FUNCTION_BLOCK PID_DEMO_PROCESS (* Offline prototype; see docs/pid/README.md; native validation pending *)
  (* Standard: 61499-2 *)
  (* Version 0.1, 2026-10-18, Guilherme *)
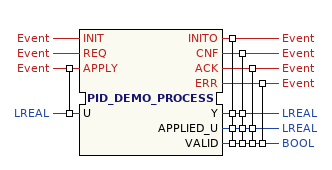
  EVENT_INPUT
    INIT;
    REQ;
    APPLY WITH U;
  END_EVENT
  EVENT_OUTPUT
    INITO WITH Y, APPLIED_U, VALID;
    CNF WITH Y, APPLIED_U, VALID;
    ACK WITH APPLIED_U, VALID;
    ERR WITH VALID;
  END_EVENT
  VAR_INPUT
    U : LREAL;
  END_VAR
  VAR_OUTPUT
    Y : LREAL;
    APPLIED_U : LREAL;
    VALID : BOOL;
  END_VAR
  VAR
    Y_NEXT : LREAL;
  END_VAR
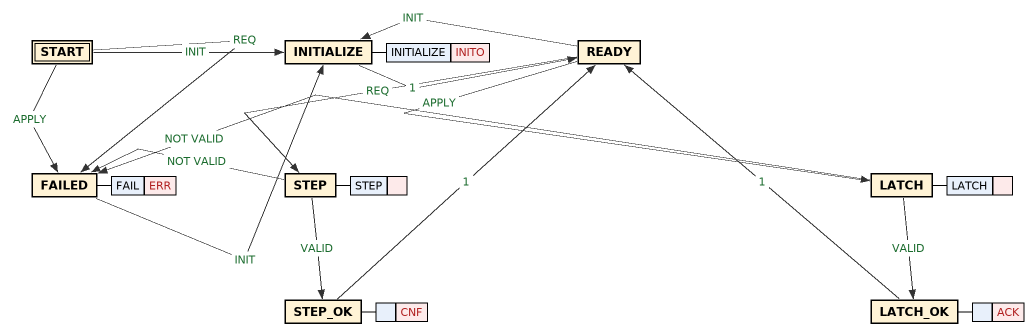
  EC_STATES
    START;
    INITIALIZE : INITIALIZE -> INITO;
    READY;
    STEP : STEP;
    STEP_OK : -> CNF;
    LATCH : LATCH;
    LATCH_OK : -> ACK;
    FAILED : FAIL -> ERR;
  END_STATES
  EC_TRANSITIONS
    START TO INITIALIZE := INIT;
    START TO FAILED := REQ;
    START TO FAILED := APPLY;
    INITIALIZE TO READY := 1;
    READY TO INITIALIZE := INIT;
    READY TO STEP := REQ;
    READY TO LATCH := APPLY;
    STEP TO STEP_OK := VALID;
    STEP TO FAILED := NOT VALID;
    STEP_OK TO READY := 1;
    LATCH TO LATCH_OK := VALID;
    LATCH TO FAILED := NOT VALID;
    LATCH_OK TO READY := 1;
    FAILED TO INITIALIZE := INIT;
  END_TRANSITIONS
  ALGORITHM INITIALIZE IN ST:
Y := 0.0;
APPLIED_U := 0.0;
VALID := TRUE;
  END_ALGORITHM
  ALGORITHM STEP IN ST:
Y_NEXT := 0.9 * Y + 0.1 * APPLIED_U;
VALID := (Y_NEXT >= -1.0E+100) AND (Y_NEXT <= 1.0E+100);
IF VALID THEN
    Y := Y_NEXT;
END_IF;
  END_ALGORITHM
  ALGORITHM LATCH IN ST:
VALID := (U >= -1.0E+100) AND (U <= 1.0E+100);
IF VALID THEN
    APPLIED_U := U;
END_IF;
  END_ALGORITHM
  ALGORITHM FAIL IN ST:
VALID := FALSE;
  END_ALGORITHM
END_FUNCTION_BLOCK
